Staubli VAL3: program.pjx

--- program.pjx ---
Parameters version=s8.15.3Cs9_BS3337 stackSize=5000 millimeterUnit=true
Program file=copy.pgx
Program file=copyItem.pgx
Program file=copyPara.pgx
Program file=deleteProg.pgx
Program file=deleteProgItem.pgx
Program file=do_CASE.pgx
Program file=do_endSwitch.pgx
Program file=do_for.pgx
Program file=do_if.pgx
Program file=do_switch.pgx
Program file=editIF.pgx
Program file=getProgItemIndex.pgx
Program file=getProgItemSize.pgx
Program file=getProgList.pgx
Program file=getSize.pgx
Program file=if_check.pgx
Program file=ifString.pgx
Program file=insertCASE.pgx
Program file=insertENDIF.pgx
Program file=insertENDSwitch.pgx
Program file=insertFOR.pgx
Program file=insertItem.pgx
Program file=insertPROG.pgx
Program file=insertSwitch.pgx
Program file=insertTRAJ.pgx
Program file=loadPROG.pgx
Program file=makeTraj.pgx
Program file=new.pgx
Program file=onSave.pgx
Program file=pointToString.pgx
Program file=start.pgx
Program file=stop.pgx
Program file=waitLoad.pgx
Data file=program.dtx
Library alias=progTemp path=Disk://source/template/progTemp/progTemp.pjx
Library alias=trajectory path=Disk://source/projectSource/trajectory/trajectory.pjx
Library alias=action path=Disk://source/projectSource/Action/Action.pjx
Library alias=rs path=Disk://source/projectSource/robotStatus/robotStatus.pjx
Library alias=io path=Disk://source/projectSource/io/io.pjx
Library alias=saveData path=Disk://source/saveData/saveData.pjx
Library alias=ar path=Disk://autoReturn/autoReturn.pjx

--- program.dtx ---
mdesc mNomSpeed
bool bError
public num nLastIndex

--- start.pgx ---
program start()
begin
end

--- copy.pgx ---
public program copy(string x_sKey, bool& x_bToSave)
  local bool l_bResult
  local string l_sName
begin
  if x_sKey!=""
    l_bResult=userPagePrompt("复制-输入新名称：",l_sName)
    if l_bResult
      if !isDefined(progTemp:pProgItem[l_sName])
        insert(progTemp:pProgItem[l_sName])
        call copyItem(l_sName,x_sKey)

        x_bToSave=true
      else
        userPageAlert("存在相同名称的程序！")
      endIf
    endIf
  endIf
end

--- copyItem.pgx ---
public program copyItem(string x_sTarget, string x_sSource)
  local num l_nSize
  local num l_i
  local num l_j
begin
  l_nSize=size(progTemp:pProgItem[x_sSource].pProgTemplate)
  resize(progTemp:pProgItem[x_sTarget].pProgTemplate,1,l_nSize)
  for l_i = 0 to l_nSize-1
    progTemp:pProgItem[x_sTarget].pProgTemplate[l_i].sTRAJname=progTemp:pProgItem[x_sSource].pProgTemplate[l_i].sTRAJname
    progTemp:pProgItem[x_sTarget].pProgTemplate[l_i].nType=progTemp:pProgItem[x_sSource].pProgTemplate[l_i].nType
    for l_j=0 to 2
      progTemp:pProgItem[x_sTarget].pProgTemplate[l_i].iIfItem.nSigType[l_j]=progTemp:pProgItem[x_sSource].pProgTemplate[l_i].iIfItem.nSigType[l_j]
      progTemp:pProgItem[x_sTarget].pProgTemplate[l_i].iIfItem.nSigIndex[l_j]=progTemp:pProgItem[x_sSource].pProgTemplate[l_i].iIfItem.nSigIndex[l_j]
      progTemp:pProgItem[x_sTarget].pProgTemplate[l_i].iIfItem.nValue[l_j]=progTemp:pProgItem[x_sSource].pProgTemplate[l_i].iIfItem.nValue[l_j]
    endFor
    progTemp:pProgItem[x_sTarget].pProgTemplate[l_i].iIfItem.bANDOR[0]=(progTemp:pProgItem[x_sSource].pProgTemplate[l_i].iIfItem.bANDOR[0]==true)
    progTemp:pProgItem[x_sTarget].pProgTemplate[l_i].iIfItem.bANDOR[1]=(progTemp:pProgItem[x_sSource].pProgTemplate[l_i].iIfItem.bANDOR[1]==true)
  endFor
end

--- copyPara.pgx ---
public program copyPara(string x_sTarget, num x_nSource, num x_nTarget)
  local num l_nSize
  local num l_i
  local num l_j
begin

  progTemp:pProgItem[x_sTarget].pProgTemplate[x_nTarget].sTRAJname=progTemp:pProgItem[x_sTarget].pProgTemplate[x_nSource].sTRAJname
  progTemp:pProgItem[x_sTarget].pProgTemplate[x_nTarget].nType=progTemp:pProgItem[x_sTarget].pProgTemplate[x_nSource].nType
  for l_j=0 to 2
    progTemp:pProgItem[x_sTarget].pProgTemplate[x_nTarget].iIfItem.nSigType[l_j]=progTemp:pProgItem[x_sTarget].pProgTemplate[x_nSource].iIfItem.nSigType[l_j]
    progTemp:pProgItem[x_sTarget].pProgTemplate[x_nTarget].iIfItem.nSigIndex[l_j]=progTemp:pProgItem[x_sTarget].pProgTemplate[x_nSource].iIfItem.nSigIndex[l_j]
    progTemp:pProgItem[x_sTarget].pProgTemplate[x_nTarget].iIfItem.nValue[l_j]=progTemp:pProgItem[x_sTarget].pProgTemplate[x_nSource].iIfItem.nValue[l_j]
  endFor
  progTemp:pProgItem[x_sTarget].pProgTemplate[x_nTarget].iIfItem.bANDOR[0]=(progTemp:pProgItem[x_sTarget].pProgTemplate[x_nSource].iIfItem.bANDOR[0]==true)
  progTemp:pProgItem[x_sTarget].pProgTemplate[x_nTarget].iIfItem.bANDOR[1]=(progTemp:pProgItem[x_sTarget].pProgTemplate[x_nSource].iIfItem.bANDOR[1]==true)

end

--- deleteProg.pgx ---
public program deleteProg(string x_sKey, bool& x_bToSave)
  local bool l_bResult
begin
  if x_sKey!=""
    l_bResult=userPageConfirm("是否删除"+x_sKey+"?")
    if l_bResult
      delete(progTemp:pProgItem[x_sKey])
      x_bToSave=true
      //progTemp:libSave()
    endIf
  endIf
end

--- deleteProgItem.pgx ---
public program deleteProgItem(string x_sKey, string x_sItem, bool& x_bToSave)
  local bool l_bResult
  local bool l_bResult1
  local num l_nIndex
begin
  if x_sItem!=""
    l_bResult=userPageConfirm("是否删除"+x_sItem+"?")
    if l_bResult
      toNum(x_sItem,l_nIndex,l_bResult1)
      if l_nIndex==0 and size(progTemp:pProgItem[x_sKey].pProgTemplate)<2
        userPageAlert("数组元素数量需大于0")
      else
        delete(progTemp:pProgItem[x_sKey].pProgTemplate[l_nIndex])
        //progTemp:libSave()
        x_bToSave=true
      endIf
    endIf
  else
    userPageAlert("未选中有效项目!")
  endIf
end

--- do_CASE.pgx ---
public program do_CASE(string x_sKey, num x_nIndex)
  local num l_nValue
  local string l_sProg
  local string l_sType
begin
  l_nValue=progTemp:pProgItem[x_sKey].pProgTemplate[x_nIndex].sSwitchItem.nSwitchValue
  l_sProg=progTemp:pProgItem[x_sKey].pProgTemplate[x_nIndex].sSwitchItem.sIOValue
  l_sType=progTemp:pProgItem[x_sKey].pProgTemplate[x_nIndex].sTRAJname
  if l_nValue==rs:nSetSwitchValue
    switch l_sType
      case "PROG"
        call makeTraj(l_sProg)
      break
      case "TRAJ"
        call trajectory:makeTraj(l_sProg)
      break
    endSwitch

    rs:nSetSwitchValue=0
    rs:bInSwitch=false
  endIf

end

--- do_endSwitch.pgx ---
public program do_endSwitch()
begin
  rs:bInSwitch=false
end

--- do_for.pgx ---
public program do_for(string x_sKey, num x_nIndex)
  local num l_nIOindex
  local bool l_bResult
  local num l_nLoop
  local bool l_bErr
  local bool l_bActive
  local string l_skey
  local num l_i
  local string l_sType
begin
  waitEndMove()
  l_bActive=false
  if progTemp:pProgItem[x_sKey].pProgTemplate[x_nIndex].fForItem.sIOindex=="value"
    l_nLoop=progTemp:pProgItem[x_sKey].pProgTemplate[x_nIndex].fForItem.nLoopValue
    l_bActive=true
  else
    toNum(progTemp:pProgItem[x_sKey].pProgTemplate[x_nIndex].fForItem.sIOindex,l_nIOindex,l_bResult)
    if l_bResult
      call io:getAnaIO(io:aInItem[l_nIOindex].aAio,l_nLoop,l_bErr)
      l_bActive=true
    endIf
  endIf
  l_skey=progTemp:pProgItem[x_sKey].pProgTemplate[x_nIndex].fForItem.sForTRAJ
  l_sType=progTemp:pProgItem[x_sKey].pProgTemplate[x_nIndex].sTRAJname
  switch l_sType
    case "PROG"
      if l_bActive
        for l_i = 0 to l_nLoop
          call makeTraj(l_skey)
        endFor
      endIf
    break
    case "TRAJ"
      if l_bActive
        for l_i = 0 to l_nLoop
          call trajectory:makeTraj(l_skey)
        endFor
      endIf
    break
  endSwitch

end

--- do_if.pgx ---
public program do_if(string x_sKey, num x_nIndex, bool& x_bResult)
  local num l_nType[3]
  local num l_nIndex[3]
  local num l_nValue[3]
  local bool l_bResult1
  local bool l_bDisable1
  local bool l_bResult2
  local bool l_bDisable2
  local bool l_bResult3
  local bool l_bDisable3
  local bool l_bANDOR1
  local bool l_bANDOR2
  local num l_i
begin
  for l_i = 0 to 2
    l_nType[l_i]=progTemp:pProgItem[x_sKey].pProgTemplate[x_nIndex].iIfItem.nSigType[l_i]
    l_nIndex[l_i]=progTemp:pProgItem[x_sKey].pProgTemplate[x_nIndex].iIfItem.nSigIndex[l_i]
    l_nValue[l_i]=progTemp:pProgItem[x_sKey].pProgTemplate[x_nIndex].iIfItem.nValue[l_i]
  endFor

  l_bANDOR1=(progTemp:pProgItem[x_sKey].pProgTemplate[x_nIndex].iIfItem.bANDOR[0]==true)
  l_bANDOR2=(progTemp:pProgItem[x_sKey].pProgTemplate[x_nIndex].iIfItem.bANDOR[1]==true)

  call if_check(l_nType[0],l_nIndex[0],l_nValue[0],l_bResult1,l_bDisable1)
  call if_check(l_nType[1],l_nIndex[1],l_nValue[1],l_bResult2,l_bDisable2)
  call if_check(l_nType[2],l_nIndex[2],l_nValue[2],l_bResult3,l_bDisable3)

  if l_bDisable2
    x_bResult=l_bResult1
  else
    if l_bANDOR1
      x_bResult=(l_bResult1 or l_bResult2)
    else
      x_bResult=(l_bResult1 and l_bResult2)
    endIf

    if l_bDisable3
    else
      if l_bANDOR2
        x_bResult=(x_bResult and (l_bResult2 or l_bResult3))
      else
        x_bResult=x_bResult and (l_bResult2 and l_bResult3)
      endIf
    endIf
  endIf



end

--- do_switch.pgx ---
public program do_switch(string x_sKey, num x_nIndex)
  local string l_sValue
  local num l_nIOindex
  local bool l_bErr
  local num l_nValue
  local bool l_bResult
begin
  waitEndMove()
  rs:bInSwitch=true
  l_sValue=progTemp:pProgItem[x_sKey].pProgTemplate[x_nIndex].sSwitchItem.sIOValue
  toNum(l_sValue,l_nIOindex,l_bResult)
  call io:getAnaIO(io:aInItem[l_nIOindex].aAio,l_nValue,l_bErr)
  rs:nSetSwitchValue=l_nValue
end

--- editIF.pgx ---
public program editIF(string x_sKey, num x_nIndex, string& x_sType[], string& x_sIOIndex[], num& x_nValue[], string x_sANDOR1, string x_sANDOR2, bool& x_bToSave)
  local num l_i
  local num l_nIndex
  local bool l_bResult
begin
  if x_nIndex==0 and progTemp:pProgItem[x_sKey].pProgTemplate[x_nIndex].sTRAJname==""
    x_nIndex=x_nIndex
  else
    x_nIndex=x_nIndex+1
    append(progTemp:pProgItem[x_sKey].pProgTemplate)
    for l_i = size(progTemp:pProgItem[x_sKey].pProgTemplate)-1 to x_nIndex step -1
      call copyPara(x_sKey,l_i-1,l_i)
    endFor
    //insert(progTemp:pProgItem[x_sKey].pProgTemplate[x_nIndex])
  endIf

  progTemp:pProgItem[x_sKey].pProgTemplate[x_nIndex].nType=3
  progTemp:pProgItem[x_sKey].pProgTemplate[x_nIndex].sTRAJname="IF"
  for l_i = 0 to 2
    if x_sIOIndex[l_i]!=""
      toNum(x_sIOIndex[l_i],l_nIndex,l_bResult)
    else
      l_nIndex=-1
    endIf
    switch x_sType[l_i]
      case "DIN"
        progTemp:pProgItem[x_sKey].pProgTemplate[x_nIndex].iIfItem.nSigType[l_i]=1
        progTemp:pProgItem[x_sKey].pProgTemplate[x_nIndex].iIfItem.nSigIndex[l_i]=l_nIndex
        progTemp:pProgItem[x_sKey].pProgTemplate[x_nIndex].iIfItem.nValue[l_i]=x_nValue[l_i]
      break
      case "DOUT"
        progTemp:pProgItem[x_sKey].pProgTemplate[x_nIndex].iIfItem.nSigType[l_i]=2
        progTemp:pProgItem[x_sKey].pProgTemplate[x_nIndex].iIfItem.nSigIndex[l_i]=l_nIndex
        progTemp:pProgItem[x_sKey].pProgTemplate[x_nIndex].iIfItem.nValue[l_i]=x_nValue[l_i]

      break
      case "AIN"
        progTemp:pProgItem[x_sKey].pProgTemplate[x_nIndex].iIfItem.nSigType[l_i]=3
        progTemp:pProgItem[x_sKey].pProgTemplate[x_nIndex].iIfItem.nSigIndex[l_i]=l_nIndex
        progTemp:pProgItem[x_sKey].pProgTemplate[x_nIndex].iIfItem.nValue[l_i]=x_nValue[l_i]

      break
      case "AOUT"
        progTemp:pProgItem[x_sKey].pProgTemplate[x_nIndex].iIfItem.nSigType[l_i]=4
        progTemp:pProgItem[x_sKey].pProgTemplate[x_nIndex].iIfItem.nSigIndex[l_i]=l_nIndex
        progTemp:pProgItem[x_sKey].pProgTemplate[x_nIndex].iIfItem.nValue[l_i]=x_nValue[l_i]

      break
      default
        progTemp:pProgItem[x_sKey].pProgTemplate[x_nIndex].iIfItem.nSigType[l_i]=0
        progTemp:pProgItem[x_sKey].pProgTemplate[x_nIndex].iIfItem.nSigIndex[l_i]=-1
        progTemp:pProgItem[x_sKey].pProgTemplate[x_nIndex].iIfItem.nValue[l_i]=0

      break
    endSwitch
  endFor

  progTemp:pProgItem[x_sKey].pProgTemplate[x_nIndex].iIfItem.bANDOR[0]=(x_sANDOR1=="OR")
  progTemp:pProgItem[x_sKey].pProgTemplate[x_nIndex].iIfItem.bANDOR[1]=(x_sANDOR2=="OR")

  x_bToSave=true
end

--- getProgItemIndex.pgx ---
public program getProgItemIndex(string x_sKey, string x_sSelProgItem, num& x_nIndex)
  local num l_nSize
  local bool l_bResult
begin
  call getProgItemSize(x_sKey,l_nSize)
  if l_nSize==1 and progTemp:pProgItem[x_sKey].pProgTemplate[0].sTRAJname==""
    x_nIndex=0
  else
    toNum(x_sSelProgItem,x_nIndex,l_bResult)
  endIf

end

--- getProgItemSize.pgx ---
public program getProgItemSize(string x_sKey, num& x_nSize)
begin
  x_nSize=size(progTemp:pProgItem[x_sKey].pProgTemplate)
end

--- getProgList.pgx ---
public program getProgList(string& x_sList[])
  local string l_sKey
begin
  resize(x_sList,1,1)
  l_sKey=first(progTemp:pProgItem)

  while l_sKey!=""
    x_sList[size(x_sList)-1]=l_sKey
    insert(x_sList[size(x_sList)])
    l_sKey=next(progTemp:pProgItem[l_sKey])
  endWhile
end

--- getSize.pgx ---
public program getSize(num& x_nSize)
begin
   if size(progTemp:pProgItem)>0
    x_nSize=size(progTemp:pProgItem)
  else
    x_nSize=1
  endIf
end

--- if_check.pgx ---
public program if_check(num x_nType, num x_nIndex, num x_nValue, bool& x_bResult, bool& x_bDisable)
  local bool l_bErr
  local bool l_bValue
  local bool l_bRecValue
  local num l_nRecValue
begin
   x_bDisable=false
    switch x_nType
      case 1
        //din
        call io:getDigIO(io:dInput[x_nIndex],l_bRecValue,l_bErr)
        l_bValue=(x_nValue!=0)
        x_bResult=(l_bRecValue==l_bValue)
      break
      case 2
        //dout
        call io:getDigIO(io:dOutput[x_nIndex],l_bRecValue,l_bErr)
        l_bValue=(x_nValue!=0)
        x_bResult=(l_bRecValue==l_bValue)
      break
      case 3
        //ain
        call io:getAnaIO(io:aInput[x_nIndex],l_nRecValue,l_bErr)
        x_bResult=(l_nRecValue==x_nValue)
      break
      case 4
        //aout
        call io:getAnaIO(io:aInput[x_nIndex],l_nRecValue,l_bErr)
        x_bResult=(l_nRecValue==x_nValue)
      break
    default
      x_bDisable=true
    break
    endSwitch

end

--- ifString.pgx ---
public program ifString(string x_sKey, num x_nIndex, string& x_sMsg)
  local num l_i
  local num l_nSigIndex
  local num l_nSigType
  local num l_nValue
  local bool l_bANDOR1
  local bool l_bANDOR2
  local string l_sMsg1
  local string l_sMsg2
  local string l_sMsg3
  local string l_sANDOR1
  local string l_sANDOR2
begin
  l_sMsg1=""
  l_sMsg2=""
  l_sMsg3=""
  l_nSigType=progTemp:pProgItem[x_sKey].pProgTemplate[x_nIndex].iIfItem.nSigType[0]
  l_nSigIndex=progTemp:pProgItem[x_sKey].pProgTemplate[x_nIndex].iIfItem.nSigIndex[0]
  l_nValue=progTemp:pProgItem[x_sKey].pProgTemplate[x_nIndex].iIfItem.nValue[0]
  if l_nSigType>0 and l_nSigIndex>0
    switch l_nSigType
      case 1
        if l_nValue!=0
          l_sMsg1="DIN"+toString("",l_nSigIndex)+"=true"
        else
          l_sMsg1="DIN"+toString("",l_nSigIndex)+"=false"
        endIf
      break
      case 2
        if l_nValue!=0
          l_sMsg1="DOUT"+toString("",l_nSigIndex)+"=true"
        else
          l_sMsg1="DOUT"+toString("",l_nSigIndex)+"=false"
        endIf
      break
      case 3
        l_sMsg1="AIN"+toString("",l_nSigIndex)+"="+toString("",l_nValue)
      break
      case 4
        l_sMsg1="AOUT"+toString("",l_nSigIndex)+"="+toString("",l_nValue)
      break
    endSwitch
  endIf
  l_bANDOR1=progTemp:pProgItem[x_sKey].pProgTemplate[x_nIndex].iIfItem.bANDOR[0]
  if !l_bANDOR1
    l_sANDOR1=" and "
  else
    l_sANDOR1=" or "
  endIf
  l_bANDOR2=progTemp:pProgItem[x_sKey].pProgTemplate[x_nIndex].iIfItem.bANDOR[1]
  if !l_bANDOR2
    l_sANDOR2=" and "
  else
    l_sANDOR2=" or "
  endIf
  l_nSigType=progTemp:pProgItem[x_sKey].pProgTemplate[x_nIndex].iIfItem.nSigType[1]
  l_nSigIndex=progTemp:pProgItem[x_sKey].pProgTemplate[x_nIndex].iIfItem.nSigIndex[1]
  l_nValue=progTemp:pProgItem[x_sKey].pProgTemplate[x_nIndex].iIfItem.nValue[1]
  if l_nSigType>0 and l_nSigIndex>0

    switch l_nSigType
      case 1
        if l_nValue!=0
          l_sMsg2="DIN"+toString("",l_nSigIndex)+"=true"
        else
          l_sMsg2="DIN"+toString("",l_nSigIndex)+"=false"
        endIf
      break
      case 2
        if l_nValue!=0
          l_sMsg2="DOUT"+toString("",l_nSigIndex)+"=true"
        else
          l_sMsg2="DOUT"+toString("",l_nSigIndex)+"=false"
        endIf
      break
      case 3
        l_sMsg2="AIN"+toString("",l_nSigIndex)+"="+toString("",l_nValue)
      break
      case 4
        l_sMsg2="AOUT"+toString("",l_nSigIndex)+"="+toString("",l_nValue)
      break
    endSwitch
    l_sMsg2=l_sANDOR1+l_sMsg2
  endIf
  l_nSigType=progTemp:pProgItem[x_sKey].pProgTemplate[x_nIndex].iIfItem.nSigType[2]
  l_nSigIndex=progTemp:pProgItem[x_sKey].pProgTemplate[x_nIndex].iIfItem.nSigIndex[2]
  l_nValue=progTemp:pProgItem[x_sKey].pProgTemplate[x_nIndex].iIfItem.nValue[2]
  if l_nSigType>0 and l_nSigIndex>0
    switch l_nSigType
      case 1
        if l_nValue!=0
          l_sMsg3="DIN"+toString("",l_nSigIndex)+"=true"
        else
          l_sMsg3="DIN"+toString("",l_nSigIndex)+"=false"
        endIf
      break
      case 2
        if l_nValue!=0
          l_sMsg3="DOUT"+toString("",l_nSigIndex)+"=true"
        else
          l_sMsg3="DOUT"+toString("",l_nSigIndex)+"=false"
        endIf
      break
      case 3
        l_sMsg3="AIN"+toString("",l_nSigIndex)+"="+toString("",l_nValue)
      break
      case 4
        l_sMsg3="AOUT"+toString("",l_nSigIndex)+"="+toString("",l_nValue)
      break
    endSwitch
    l_sMsg3=l_sANDOR2+l_sMsg3
  endIf

  x_sMsg=l_sMsg1+l_sMsg2+l_sMsg3
end

--- insertCASE.pgx ---
public program insertCASE(string x_sKey, num x_nIndex, string x_sTRAJname, bool& x_bToSave, num x_nSwitchValue, num x_nType)
  local num l_nIndex
  local num l_i
begin

  if x_nIndex==0 and progTemp:pProgItem[x_sKey].pProgTemplate[x_nIndex].sTRAJname==""
    progTemp:pProgItem[x_sKey].pProgTemplate[x_nIndex].nType=6
    if x_nType==1
      progTemp:pProgItem[x_sKey].pProgTemplate[x_nIndex].sTRAJname="PROG"
    elseIf x_nType==2
      progTemp:pProgItem[x_sKey].pProgTemplate[x_nIndex].sTRAJname="TRAJ"
    endIf
    progTemp:pProgItem[x_sKey].pProgTemplate[x_nIndex].sSwitchItem.sIOValue=x_sTRAJname
    progTemp:pProgItem[x_sKey].pProgTemplate[x_nIndex].sSwitchItem.nSwitchValue=x_nSwitchValue
  else
    l_nIndex=x_nIndex+1
    //insert(progTemp:pProgItem[x_sKey].pProgTemplate[x_nIndex+1])
    append(progTemp:pProgItem[x_sKey].pProgTemplate)
    for l_i = size(progTemp:pProgItem[x_sKey].pProgTemplate)-1 to l_nIndex step -1
      call copyPara(x_sKey,l_i-1,l_i)
    endFor
    //insert(progTemp:pProgItem[x_sKey].pProgTemplate[x_nIndex+1])
    progTemp:pProgItem[x_sKey].pProgTemplate[x_nIndex+1].nType=6
    if x_nType==1
      progTemp:pProgItem[x_sKey].pProgTemplate[x_nIndex+1].sTRAJname="PROG"
    elseIf x_nType==2
      progTemp:pProgItem[x_sKey].pProgTemplate[x_nIndex+1].sTRAJname="TRAJ"
    endIf
    progTemp:pProgItem[x_sKey].pProgTemplate[x_nIndex+1].sSwitchItem.sIOValue=x_sTRAJname
    progTemp:pProgItem[x_sKey].pProgTemplate[x_nIndex+1].sSwitchItem.nSwitchValue=x_nSwitchValue
  endIf

  x_bToSave=true
end

--- insertENDIF.pgx ---
public program insertENDIF(string x_sKey, num x_nIndex, bool& x_bToSave)
  local num l_i
begin
  if x_nIndex==0 and progTemp:pProgItem[x_sKey].pProgTemplate[x_nIndex].sTRAJname==""
    x_nIndex=x_nIndex
  else
    x_nIndex=x_nIndex+1
    //insert(progTemp:pProgItem[x_sKey].pProgTemplate[x_nIndex])
     //l_nIndex=x_nIndex+1
    //insert(progTemp:pProgItem[x_sKey].pProgTemplate[x_nIndex+1])
    append(progTemp:pProgItem[x_sKey].pProgTemplate)
    for l_i = size(progTemp:pProgItem[x_sKey].pProgTemplate)-1 to x_nIndex step -1
      call copyPara(x_sKey,l_i-1,l_i)
    endFor
  endIf

  progTemp:pProgItem[x_sKey].pProgTemplate[x_nIndex].nType=4
  progTemp:pProgItem[x_sKey].pProgTemplate[x_nIndex].sTRAJname="ENDIF"
  x_bToSave=true
end

--- insertENDSwitch.pgx ---
public program insertENDSwitch(string x_sKey, num x_nIndex, bool& x_bToSave)
  local num l_i
begin
  if x_nIndex==0 and progTemp:pProgItem[x_sKey].pProgTemplate[x_nIndex].sTRAJname==""
    x_nIndex=x_nIndex
  else
    x_nIndex=x_nIndex+1
    //// insert(progTemp:pProgItem[x_sKey].pProgTemplate[x_nIndex])
    //l_nIndex=x_nIndex+1
    //insert(progTemp:pProgItem[x_sKey].pProgTemplate[x_nIndex+1])
    append(progTemp:pProgItem[x_sKey].pProgTemplate)
    for l_i = size(progTemp:pProgItem[x_sKey].pProgTemplate)-1 to x_nIndex step -1
      call copyPara(x_sKey,l_i-1,l_i)
    endFor
  endIf

  progTemp:pProgItem[x_sKey].pProgTemplate[x_nIndex].nType=7
  progTemp:pProgItem[x_sKey].pProgTemplate[x_nIndex].sTRAJname="ENDSWITCH"
  x_bToSave=true
end

--- insertFOR.pgx ---
public program insertFOR(string x_sKey, num x_nIndex, string x_sTRAJname, num x_nLoop, string x_sIOindex, bool x_bToSave, num x_nType)
  local num l_nIndex
  local num l_i
begin

  if x_nIndex==0 and progTemp:pProgItem[x_sKey].pProgTemplate[x_nIndex].sTRAJname==""
    progTemp:pProgItem[x_sKey].pProgTemplate[x_nIndex].nType=8
    if x_nType==1
      progTemp:pProgItem[x_sKey].pProgTemplate[x_nIndex].sTRAJname="PROG"
    elseIf x_nType==2
      progTemp:pProgItem[x_sKey].pProgTemplate[x_nIndex].sTRAJname="TRAJ"
    endIf
    progTemp:pProgItem[x_sKey].pProgTemplate[x_nIndex].fForItem.sForTRAJ=x_sTRAJname
    progTemp:pProgItem[x_sKey].pProgTemplate[x_nIndex].fForItem.nLoopValue=x_nLoop
    progTemp:pProgItem[x_sKey].pProgTemplate[x_nIndex].fForItem.sIOindex=x_sIOindex
  else
    //insert(progTemp:pProgItem[x_sKey].pProgTemplate[x_nIndex+1])
    l_nIndex=x_nIndex+1
    //insert(progTemp:pProgItem[x_sKey].pProgTemplate[x_nIndex+1])
    append(progTemp:pProgItem[x_sKey].pProgTemplate)
    for l_i = size(progTemp:pProgItem[x_sKey].pProgTemplate)-1 to l_nIndex step -1
      call copyPara(x_sKey,l_i-1,l_i)
    endFor
    progTemp:pProgItem[x_sKey].pProgTemplate[x_nIndex+1].nType=8
    if x_nType==1
      progTemp:pProgItem[x_sKey].pProgTemplate[x_nIndex+1].sTRAJname="PROG"
    elseIf x_nType==2
      progTemp:pProgItem[x_sKey].pProgTemplate[x_nIndex+1].sTRAJname="TRAJ"
    endIf
    progTemp:pProgItem[x_sKey].pProgTemplate[x_nIndex+1].fForItem.sForTRAJ=x_sTRAJname
    progTemp:pProgItem[x_sKey].pProgTemplate[x_nIndex+1].fForItem.nLoopValue=x_nLoop
    progTemp:pProgItem[x_sKey].pProgTemplate[x_nIndex+1].fForItem.sIOindex=x_sIOindex
  endIf

  x_bToSave=true
end

--- insertItem.pgx ---
public program insertItem(string x_sKey, string& x_sIndex, string x_sTRAJname, num x_nType, bool& x_bToSave)
  local num l_nIndex
  local bool l_bResult
  local num l_i
begin
  if x_sIndex!=""
    toNum(x_sIndex,l_nIndex,l_bResult)
    if l_bResult
      if l_nIndex==0 and progTemp:pProgItem[x_sKey].pProgTemplate[l_nIndex].sTRAJname==""
        progTemp:pProgItem[x_sKey].pProgTemplate[l_nIndex].sTRAJname=x_sTRAJname
        progTemp:pProgItem[x_sKey].pProgTemplate[l_nIndex].nType=x_nType
      else
        // l_nIndex=l_nIndex+1
        //insert(progTemp:pProgItem[x_sKey].pProgTemplate[l_nIndex])
        //l_nIndex=x_nIndex+1
        //insert(progTemp:pProgItem[x_sKey].pProgTemplate[x_nIndex+1])
        append(progTemp:pProgItem[x_sKey].pProgTemplate)
        for l_i = size(progTemp:pProgItem[x_sKey].pProgTemplate)-1 to l_nIndex step -1
          call copyPara(x_sKey,l_i-1,l_i)
        endFor
        progTemp:pProgItem[x_sKey].pProgTemplate[l_nIndex].sTRAJname=x_sTRAJname
        progTemp:pProgItem[x_sKey].pProgTemplate[l_nIndex].nType=x_nType
      endIf
      switch x_nType
        case 0
          x_sIndex=toString("",l_nIndex)+",TRAJ->"+x_sTRAJname
        break
        case 1
          x_sIndex=toString("",l_nIndex)+",ACTION->"+x_sTRAJname
        break
        case 2
          x_sIndex=toString("",l_nIndex)+",PROG->"+x_sTRAJname
        break
      endSwitch

      x_bToSave=true
    endIf
  else
    userPageAlert("未选中项目！")
  endIf
end

--- insertPROG.pgx ---
public program insertPROG(string x_sKey, num x_nIndex, string x_sTRAJname, bool& x_bToSave)
  local num l_nIndex
  local num l_i
begin
  if x_nIndex==0 and progTemp:pProgItem[x_sKey].pProgTemplate[x_nIndex].sTRAJname==""
    progTemp:pProgItem[x_sKey].pProgTemplate[x_nIndex].nType=2
    progTemp:pProgItem[x_sKey].pProgTemplate[x_nIndex].sTRAJname=x_sTRAJname
  else
    //insert(progTemp:pProgItem[x_sKey].pProgTemplate[x_nIndex+1])
    l_nIndex=x_nIndex+1
    //insert(progTemp:pProgItem[x_sKey].pProgTemplate[x_nIndex+1])
    append(progTemp:pProgItem[x_sKey].pProgTemplate)
    for l_i = size(progTemp:pProgItem[x_sKey].pProgTemplate)-1 to l_nIndex step -1
      call copyPara(x_sKey,l_i-1,l_i)
    endFor
    progTemp:pProgItem[x_sKey].pProgTemplate[x_nIndex+1].nType=2
    progTemp:pProgItem[x_sKey].pProgTemplate[x_nIndex+1].sTRAJname=x_sTRAJname
  endIf

  x_bToSave=true
end

--- insertSwitch.pgx ---
public program insertSwitch(string x_sKey, num x_nIndex, string x_sValue, bool x_bToSave)
  local num l_i
begin
  if x_nIndex==0 and progTemp:pProgItem[x_sKey].pProgTemplate[x_nIndex].sTRAJname==""
    x_nIndex=x_nIndex
  else
    x_nIndex=x_nIndex+1
    //insert(progTemp:pProgItem[x_sKey].pProgTemplate[x_nIndex])
    //l_nIndex=x_nIndex+1
    //insert(progTemp:pProgItem[x_sKey].pProgTemplate[x_nIndex+1])
    append(progTemp:pProgItem[x_sKey].pProgTemplate)
    for l_i = size(progTemp:pProgItem[x_sKey].pProgTemplate)-1 to x_nIndex step -1
      call copyPara(x_sKey,l_i-1,l_i)
    endFor
  endIf

  progTemp:pProgItem[x_sKey].pProgTemplate[x_nIndex].nType=5
  progTemp:pProgItem[x_sKey].pProgTemplate[x_nIndex].sTRAJname="SWITCH"
  progTemp:pProgItem[x_sKey].pProgTemplate[x_nIndex].sSwitchItem.sIOValue=x_sValue
  progTemp:pProgItem[x_sKey].pProgTemplate[x_nIndex].sSwitchItem.bIOdisable=true
  //insert(progTemp:pProgItem[x_sKey].pProgTemplate[x_nIndex+1])
  append(progTemp:pProgItem[x_sKey].pProgTemplate)
  for l_i = size(progTemp:pProgItem[x_sKey].pProgTemplate)-1 to(x_nIndex+1) step -1
    call copyPara(x_sKey,l_i-1,l_i)
  endFor
  progTemp:pProgItem[x_sKey].pProgTemplate[x_nIndex+1].nType=7
  progTemp:pProgItem[x_sKey].pProgTemplate[x_nIndex+1].sTRAJname="ENDSWITCH"
  //progTemp:pProgItem[x_sKey].pProgTemplate[x_nIndex].sSwitchItem.sIOValue=x_nValue
  //progTemp:pProgItem[x_sKey].pProgTemplate[x_nIndex].sSwitchItem.bIOdisable=true

  x_bToSave=true
end

--- insertTRAJ.pgx ---
public program insertTRAJ(string x_sKey, num x_nIndex, string x_sTRAJname, bool& x_bToSave)
  local num l_nIndex
  local num l_i
begin
  if x_nIndex==0 and progTemp:pProgItem[x_sKey].pProgTemplate[x_nIndex].sTRAJname==""
    progTemp:pProgItem[x_sKey].pProgTemplate[x_nIndex].nType=0
    progTemp:pProgItem[x_sKey].pProgTemplate[x_nIndex].sTRAJname=x_sTRAJname
  else
    l_nIndex=x_nIndex+1
    //insert(progTemp:pProgItem[x_sKey].pProgTemplate[x_nIndex+1])
    append(progTemp:pProgItem[x_sKey].pProgTemplate)
    for l_i = size(progTemp:pProgItem[x_sKey].pProgTemplate)-1 to l_nIndex step -1
      call copyPara(x_sKey,l_i-1,l_i)
    endFor
    progTemp:pProgItem[x_sKey].pProgTemplate[x_nIndex+1].nType=0
    progTemp:pProgItem[x_sKey].pProgTemplate[x_nIndex+1].sTRAJname=x_sTRAJname
  endIf

  x_bToSave=true
end

--- loadPROG.pgx ---
public program loadPROG(num x_nLib, num& x_nResult)
  local string l_sPath
  local num l_nClock
begin
  l_nClock=clock()
  if x_nLib>=0

    l_sPath="Disk://data/CustomerLib/lib"+toString("",x_nLib)+"/savePROG"
    x_nResult=progTemp:libLoad(l_sPath)
    if x_nResult!=0
      popUpMsg("1")
      call rs:setAlarm(300,0)
    endIf
  else
    call rs:setAlarm(302,0)
  endIf
  logMsg(progTemp:libPath()+",耗时:"+toString(".3",clock()-l_nClock))

end

--- makeTraj.pgx ---
public program makeTraj(string x_sKey)
  local string l_sType
  local string l_sTrajName
  local num l_i
  local num l_nIndex
  local bool l_bResult
  local num l_nType
  local num l_nResult
begin
  //  if nLastIndex!=saveData:nLibIndex
  //    nLastIndex=saveData:nLibIndex
  //    call loadPROG(saveData:nLibIndex,l_nResult)
  //    call trajectory:loadTRAJ(saveData:nLibIndex,l_nResult)
  //    delay(1)
  //  endIf
  call ar:resetReturnStack(false)
  if isDefined(progTemp:pProgItem[x_sKey])
    // rs:bProgGOTO=false
    for l_i = 0 to size(progTemp:pProgItem[x_sKey].pProgTemplate)-1
      l_nType=progTemp:pProgItem[x_sKey].pProgTemplate[l_i].nType
      l_sTrajName=progTemp:pProgItem[x_sKey].pProgTemplate[l_i].sTRAJname
      if !rs:bProgGOTO
        switch l_nType
          case 0
            call trajectory:makeTraj(l_sTrajName)
          break
          case 1
            toNum(l_sTrajName,l_nIndex,l_bResult)
            call action:action_do(l_nIndex)
          break
          case 2
            call makeTraj(l_sTrajName)
          break
          case 3
            waitEndMove()
            call do_if(x_sKey,l_i,l_bResult)
            rs:bProgGOTO=(l_bResult==false)
          break
          case 4
            waitEndMove()
            rs:bProgGOTO=false
          break
          case 5
            call do_switch(x_sKey,l_i)
          break
          case 6
            call do_CASE(x_sKey,l_i)
          break
          case 7
            call do_endSwitch()
          break
          case 8
            call do_for(x_sKey,l_i)
          break

        endSwitch
      else
        if l_nType==4
          rs:bProgGOTO=false
        endIf
      endIf
      delay(0)
    endFor
  else
    bError=true
    popUpMsg("program:"+x_sKey+" 未定义")
  endIf
  waitEndMove()
end

--- new.pgx ---
public program new(bool& x_bToSave)
  local string l_sNmae
  local bool l_bResult
begin
  l_bResult=userPagePrompt("输入新建名称：",l_sNmae)
  if l_bResult
    if !isDefined(progTemp:pProgItem[l_sNmae])
      insert(progTemp:pProgItem[l_sNmae])
      x_bToSave=true
    endIf
  endIf
end

--- onSave.pgx ---
public program onSave(bool& x_bTosave)
begin
  if x_bTosave
    rs:bIsSaving=true
    progTemp:libSave()
    x_bTosave=false
    rs:bIsSaving=false
    delay(0.1)
    popUpMsg("数据已保存")
  endIf
end

--- pointToString.pgx ---
public program pointToString(string& x_sMsg, string x_sKey, num x_nIndex)
  local string l_sMsg
  local num l_nType
  local string l_sType
  local string l_sMsg1
  local string l_sTrajName
  local string l_sType1
begin
  l_nType=progTemp:pProgItem[x_sKey].pProgTemplate[x_nIndex].nType
  l_sTrajName=progTemp:pProgItem[x_sKey].pProgTemplate[x_nIndex].sTRAJname
  if l_sTrajName!=""
    switch l_nType
      case 0
        l_sType="TRAJ"
      break
      case 1
        l_sType="ACTION"
      break
      case 2
        l_sType="PROG"
      break
      case 3
        l_sType="IF"
      break
      case 4
        l_sType="ENDIF"
      break
      case 5
        l_sType="SWITCH"
      break
      case 6
        l_sType="---CASE"
      break
      case 7
        l_sType="ENDSWITCH"
      break
      case 8
        l_sType="FOR"
      break
      default
      break
    endSwitch
    if l_nType<3
      l_sMsg=" |"
      l_sMsg=l_sMsg+l_sType
      l_sMsg=l_sMsg+" -> "+progTemp:pProgItem[x_sKey].pProgTemplate[x_nIndex].sTRAJname
      x_sMsg=l_sMsg
    elseIf l_nType==3
      call ifString(x_sKey,x_nIndex,l_sMsg1)
      l_sMsg=" |IF "
      l_sMsg=l_sMsg+l_sMsg1
      x_sMsg=l_sMsg
    elseIf l_nType==4
      l_sMsg=" |"
      l_sMsg=l_sMsg+"ENDIF"
      x_sMsg=l_sMsg
    elseIf l_nType==5
      l_sMsg=" |"
      l_sMsg=l_sMsg+l_sType+" ["+progTemp:pProgItem[x_sKey].pProgTemplate[x_nIndex].sSwitchItem.sIOValue+"]"
      x_sMsg=l_sMsg
    elseIf l_nType==7
      l_sMsg=" |"+l_sType
      x_sMsg=l_sMsg
    elseIf l_nType==6
      l_sType1=progTemp:pProgItem[x_sKey].pProgTemplate[x_nIndex].sTRAJname
      l_sMsg=" |"+l_sType+"  "+toString("",progTemp:pProgItem[x_sKey].pProgTemplate[x_nIndex].sSwitchItem.nSwitchValue)
      l_sMsg=l_sMsg+" -> "+l_sType1+" ["+progTemp:pProgItem[x_sKey].pProgTemplate[x_nIndex].sSwitchItem.sIOValue+"]"
      x_sMsg=l_sMsg
    elseIf l_nType==8
      if progTemp:pProgItem[x_sKey].pProgTemplate[x_nIndex].fForItem.sIOindex=="value"
        l_sMsg=" |"+l_sType+" to [value="+toString("",progTemp:pProgItem[x_sKey].pProgTemplate[x_nIndex].fForItem.nLoopValue)+"]"
      else
        l_sMsg=" |"+l_sType+" to AIN｛"+progTemp:pProgItem[x_sKey].pProgTemplate[x_nIndex].fForItem.sIOindex+"｝"
      endIf
      l_sMsg=l_sMsg+" -> "+progTemp:pProgItem[x_sKey].pProgTemplate[x_nIndex].fForItem.sForTRAJ
      x_sMsg=l_sMsg
    endIf
  endIf
end

--- stop.pgx ---
program stop()
begin
end

--- waitLoad.pgx ---
public program waitLoad(num x_nLib)
  local string l_sPath
  local string l_sPath1
begin
  l_sPath="Disk://data/CustomerLib/lib"+toString("",x_nLib)+"/savePROG"

  do
    l_sPath1=progTemp:libPath()
    delay(0)
  until l_sPath==l_sPath1
end
